TYPE ET_ItpReadRParams :
(
	ET_ItpReadRParams_eWaitExecute := 0,
	ET_ItpReadRParams_eReadRParams := 5,
	ET_ItpReadRParams_eDone := 197,
	ET_ItpReadRParams_eError := 198,
	ET_ItpReadRParams_eNoExecute := 199
);
END_TYPE

(* stored: Version 1.1.0.1, ProductVersion 3.1.4024.15
   DUT ET_ItpReadRParams: Id {5867cf5d-08a2-4a85-a420-d5cd034ebec7} *)
